// TIA Portal V18 export
TYPE "InterlockEmergMdz_in"
   STRUCT
      StationInterlock_APLC_Input : Array[1.."Station_Setup_Const"] of Struct
         Emergencial_Interlock_APLC_Input : Bool;
      END_STRUCT;
   END_STRUCT;
END_TYPE
